% RSLogix 500 project PROGRAM 9.RSS, saved by version 8.30.00.16 %
PROJECT "UNTITLED"    % processor: Bul.1763 MicroLogix 1100 Series B %

PROGRAM FILES
  LAD 2 "MAIN"  2 rungs
  LAD 3 "IO"  8 rungs

DATA FILES
  O0 OUTPUT  4 elements
  I1 INPUT  6 elements
  S2 STATUS  66 elements
  B3 BINARY  1 elements
  T4 TIMER  1 elements
  C5 COUNTER  1 elements
  R6 CONTROL  1 elements
  N7 INTEGER  4 elements
  F8 FLOAT  1 elements
  ST9   3 elements
  ST10   4 elements

LADDER 2 "MAIN"
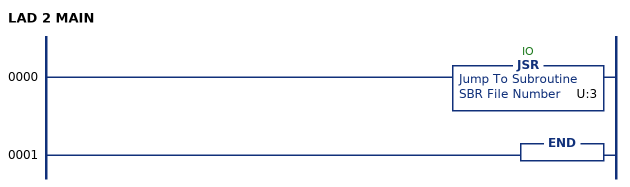
% Rung: 0 %
SOR JSR U:3 EOR
%   U:3  "IO" %
% Rung: 1 %
SOR END EOR

LADDER 3 "IO"
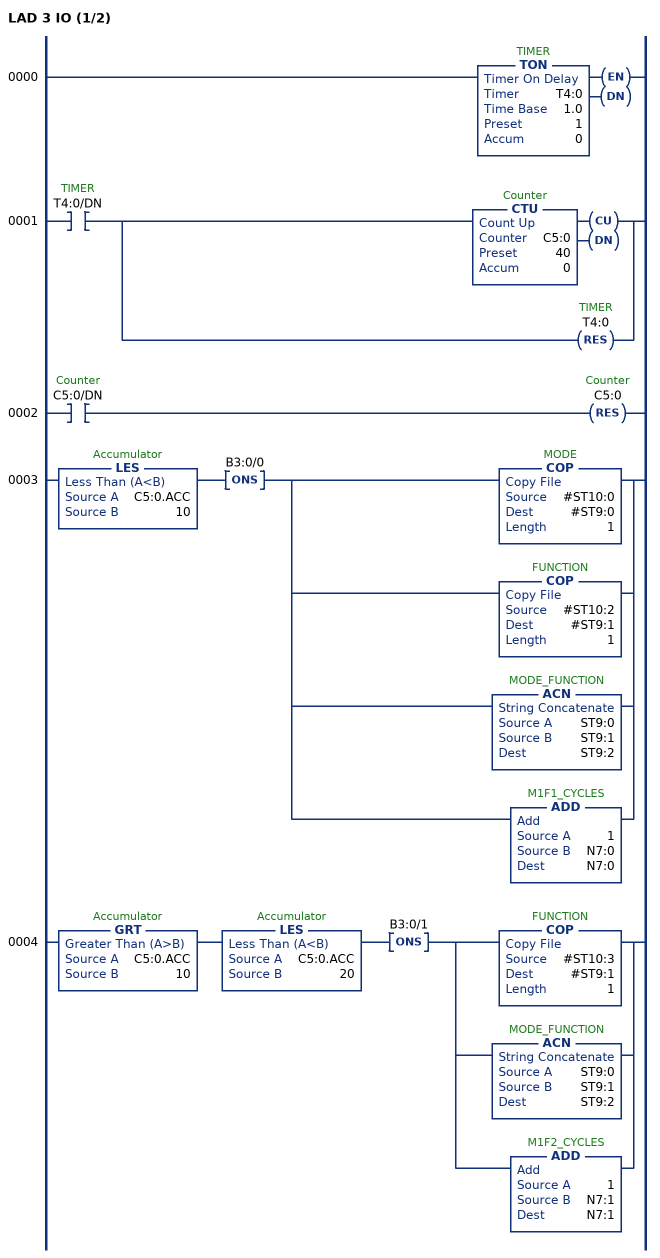
% Rung: 0 %
SOR TON T4:0 1.0 1 0 EOR
%   T4:0  "TIMER" %
% Rung: 1 %
SOR XIC T4:0/DN BST CTU C5:0 40 0 NXB RES T4:0 BND EOR
%   T4:0  "TIMER" %
%   C5:0  "Counter" %
% Rung: 2 %
SOR XIC C5:0/DN RES C5:0 EOR
%   C5:0  "Counter" %
% Rung: 3 %
SOR LES C5:0.ACC 10 ONS B3:0/0 BST COP #ST10:0 #ST9:0 1 NXB COP #ST10:2 #ST9:1 1 NXB ACN ST9:0 ST9:1 ST9:2 NXB ADD 1 N7:0 N7:0 BND EOR
%   C5:0.ACC  "Accumulator" %
%   ST9:0  MODE %
%   ST9:1  FUNCTION %
%   ST9:2  MODE_FUNCTION %
%   N7:0  M1F1_CYCLES %
% Rung: 4 %
SOR GRT C5:0.ACC 10 LES C5:0.ACC 20 ONS B3:0/1 BST COP #ST10:3 #ST9:1 1 NXB ACN ST9:0 ST9:1 ST9:2 NXB ADD 1 N7:1 N7:1 BND EOR
%   C5:0.ACC  "Accumulator" %
%   ST9:1  FUNCTION %
%   ST9:0  MODE %
%   ST9:2  MODE_FUNCTION %
%   N7:1  M1F2_CYCLES %

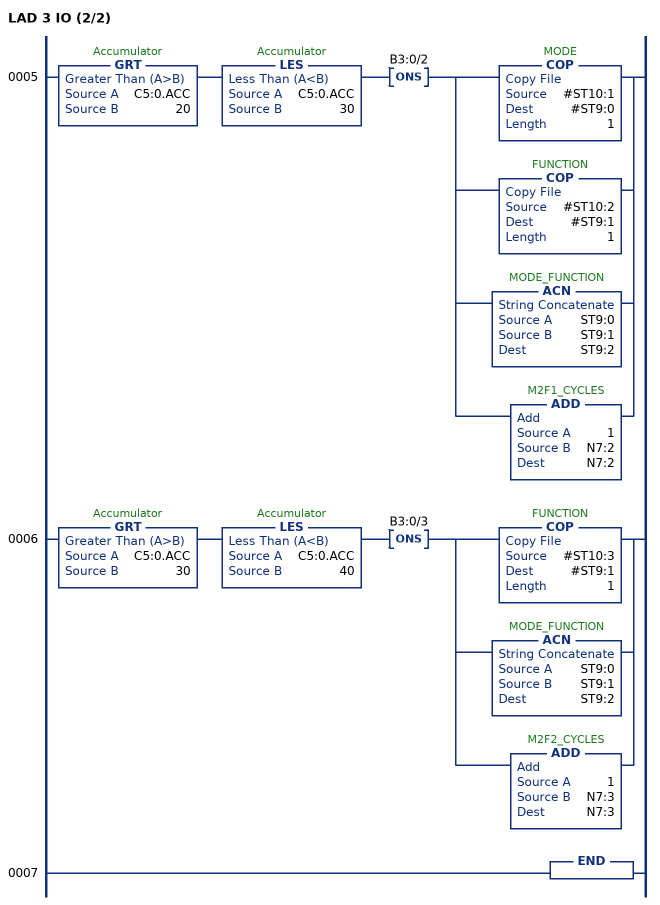
% Rung: 5 %
SOR GRT C5:0.ACC 20 LES C5:0.ACC 30 ONS B3:0/2 BST COP #ST10:1 #ST9:0 1 NXB COP #ST10:2 #ST9:1 1 NXB ACN ST9:0 ST9:1 ST9:2 NXB ADD 1 N7:2 N7:2 BND EOR
%   C5:0.ACC  "Accumulator" %
%   ST9:0  MODE %
%   ST9:1  FUNCTION %
%   ST9:2  MODE_FUNCTION %
%   N7:2  M2F1_CYCLES %
% Rung: 6 %
SOR GRT C5:0.ACC 30 LES C5:0.ACC 40 ONS B3:0/3 BST COP #ST10:3 #ST9:1 1 NXB ACN ST9:0 ST9:1 ST9:2 NXB ADD 1 N7:3 N7:3 BND EOR
%   C5:0.ACC  "Accumulator" %
%   ST9:1  FUNCTION %
%   ST9:0  MODE %
%   ST9:2  MODE_FUNCTION %
%   N7:3  M2F2_CYCLES %
% Rung: 7 %
SOR END EOR

OTHER DOCUMENTED ADDRESSES
  B3:0  "ONS"
  B3:1  "ONS"
  B3:2  "ONS"
  B3:3  "ONS"
  B3:4  "ONS"
  CT54:0  "Counter"

DATA TABLE (non-zero values as saved)
DATA T4
% .PRE .ACC %
% T4:0 % 1 0
DATA C5
% .PRE .ACC %
% C5:0 % 40 0
DATA ST10
% ST10:0 % "MODE_1"
% ST10:1 % "MODE_2"
% ST10:2 % "FUNCTION_1"
% ST10:3 % "FUNCTION_2"
